// TIA Portal V21 export
Screen "R08_Sym"  1024x768, Number=48, Template=Tpl
  ScreenLayer 
    SymbolicIOField "P_SymIO" at 10,10 size 100x30  Mode=Output, TextList=TL_State
      ProcessValue := P_Cell
